// TIA Portal V20 export
TYPE "Eingänge_Zählerbaugruppe"
   STRUCT
      "COUNT VALUE" : DInt;   // Aktueller Zählwert
      "CAPTURED VALUE" : DInt;   // Letzter erfasster Capture-Wert
      "MEASURED VALUE" : DInt;   // Aktueller Messwert
      POWER_ERROR : Bool;   // Bit 0: Fehlerhafte Versorgungsspannung L+
      ENC_ERROR : Bool;   // Bit 1: Fehlerhaftes Gebersignal
      LD_ERROR : Bool;   // Bit 2: Fehler beim Laden über Steuerschnittstelle
      Reserve : Bool;   // Bit 3 bis 7: Reserve; auf 0 gesetzt
      Reserve_1 : Bool;
      Reserve_2 : Bool;
      Reserve_3 : Bool;
      Reserve_4 : Bool;
      Reserve_t : Bool;   // Bit 0: Reserve; auf 0 gesetzt
      RES_EVENT_ACK : Bool;   // Bit 1: Rücksetzen der Statusbits aktiv
      LD_STS_SLOT_0 : Bool;   // Bit 2: Ladeaufforderung für Slot 0 erkannt und durchgeführt (toggelnd)
      LD_STS_SLOT_1 : Bool;   // Bit 3: Ladeaufforderung für Slot 1 erkannt und durchgeführt (toggelnd)
      STS_READY : Bool;   // Bit 4: Technologiemodul angelaufen und parametriert
      STS_SW_GATE : Bool;   // Bit 5: Zustand SW-Tor
      Reserve_z : Bool;   // Bit 6 bis 7: Reserve; auf 0 gesetzt
      Reserve_z_1 : Bool;
      STS_DIR : Bool;   // Bit 0: Richtung der letzten Zählwertänderung
      STS_CNT : Bool;   // Bit 1: Zählimpuls innerhalb der letzten 0,5 s erfasst
      STS_GATE : Bool;   // Bit 2: Zustand internes Tor
      STS_DQ0 : Bool;   // Bit 3: Zustand DQ0
      STS_DQ1 : Bool;   // Bit 4: Zustand DQ1
      STS_DI0 : Bool;   // Bit 5: Zustand DI0
      STS_DI1 : Bool;   // Bit 6: Zustand DI1
      STS_DI2 : Bool;   // Bit 7: Zustand DI2
      EVENT_ZERO : Bool;   // Bit 0: Nulldurchgang aufgetreten
      EVENT_UFLW : Bool;   // Bit 1: Unterlauf aufgetreten
      EVENT_OFLW : Bool;   // Bit 2: Überlauf aufgetreten
      EVENT_CMP0 : Bool;   // Bit 3: Vergleichsereignis für DQ0 aufgetreten
      EVENT_CMP1 : Bool;   // Bit 4: Vergleichsereignis für DQ1 aufgetreten
      EVENT_SYNC : Bool;   // Bit 5: Synchronisation aufgetreten
      EVENT_CAP : Bool;   // Bit 6: Capture-Ereignis aufgetreten
      STS_M_INTERVAL : Bool;   // Bit 7: Zählimpuls im vorangegangenen Messintervall erfasst
   END_STRUCT;
END_TYPE
